(* IEC 61131-3 sources: llm-plc-st-eval/data/processed_definitivo/gpt-4o-2024-08-06/A4/few_shot, 3 files *)

(* ---- ejec_1.st ---- *)
FUNCTION_BLOCK FB_Rampa
VAR_INPUT
    SPvel : REAL; (* Consigna de velocidad *)
    paroRapido : BOOL; (* Activar paro rápido *)
    ciclo : TIME; (* Período de ejecución del bloque *)
END_VAR
VAR_OUTPUT
    CVvel : REAL; (* Velocidad de consigna con rampa *)
END_VAR
VAR
    incremento : REAL; (* Incremento calculado por ciclo *)
    tiempoSegundos : REAL; (* Tiempo de ciclo en segundos *)
END_VAR

(* Convertir el tiempo de ciclo a segundos *)
tiempoSegundos := REAL_TO_REAL(TIME_TO_REAL(ciclo)) / 1000.0;

IF paroRapido THEN
    (* Paro rápido: disminuir CVvel hacia 0.0 con pendiente de 40.0 puntos porcentuales por segundo *)
    incremento := -40.0 * tiempoSegundos;
    CVvel := CVvel + incremento;
    IF CVvel < 0.0 THEN
        CVvel := 0.0;
    END_IF
ELSE
    (* Ajuste normal de CVvel hacia SPvel *)
    IF SPvel > CVvel THEN
        (* Aumentar CVvel hacia SPvel con pendiente de 10.0 puntos porcentuales por segundo *)
        incremento := 10.0 * tiempoSegundos;
        CVvel := CVvel + incremento;
        IF CVvel > SPvel THEN
            CVvel := SPvel;
        END_IF
    ELSIF SPvel < CVvel THEN
        (* Disminuir CVvel hacia SPvel con pendiente de 20.0 puntos porcentuales por segundo *)
        incremento := -20.0 * tiempoSegundos;
        CVvel := CVvel + incremento;
        IF CVvel < SPvel THEN
            CVvel := SPvel;
        END_IF
    END_IF
END_IF
END_FUNCTION_BLOCK

(* ---- ejec_2.st ---- *)
FUNCTION_BLOCK FB_Rampa
VAR_INPUT
    SPvel : REAL; (* Consigna de velocidad *)
    paroRapido : BOOL; (* Señal de paro rápido *)
    ciclo : TIME; (* Período de ejecución del bloque *)
END_VAR
VAR_OUTPUT
    CVvel : REAL; (* Velocidad de consigna con rampa *)
END_VAR
VAR
    incremento : REAL; (* Incremento de velocidad por ciclo *)
    tiempoSegundos : REAL; (* Duración del ciclo en segundos *)
END_VAR

(* Convertir el tiempo de ciclo a segundos *)
tiempoSegundos := REAL_TO_REAL(TIME_TO_REAL(ciclo)) / 1000.0;

IF paroRapido THEN
    (* Paro rápido: disminuir CVvel a 0.0 con pendiente de 40.0 %/s *)
    incremento := -40.0 * tiempoSegundos;
    CVvel := CVvel + incremento;
    IF CVvel < 0.0 THEN
        CVvel := 0.0;
    END_IF
ELSE
    (* Rampa normal: ajustar CVvel hacia SPvel *)
    IF SPvel > CVvel THEN
        (* Incremento al subir con pendiente de 10.0 %/s *)
        incremento := 10.0 * tiempoSegundos;
        CVvel := CVvel + incremento;
        IF CVvel > SPvel THEN
            CVvel := SPvel;
        END_IF
    ELSIF SPvel < CVvel THEN
        (* Decremento al bajar con pendiente de 20.0 %/s *)
        incremento := -20.0 * tiempoSegundos;
        CVvel := CVvel + incremento;
        IF CVvel < SPvel THEN
            CVvel := SPvel;
        END_IF
    END_IF
END_IF
END_FUNCTION_BLOCK

(* ---- ejec_3.st ---- *)
FUNCTION_BLOCK FB_Rampa
VAR_INPUT
    SPvel : REAL; (* Consigna de velocidad *)
    paroRapido : BOOL; (* Señal de paro rápido *)
    ciclo : TIME; (* Período de ejecución del bloque *)
END_VAR
VAR_OUTPUT
    CVvel : REAL; (* Velocidad de consigna con rampa *)
END_VAR
VAR
    deltaTiempo : REAL; (* Tiempo de ciclo en segundos *)
    incremento : REAL; (* Incremento de velocidad por ciclo *)
END_VAR

(* Convertir el tiempo de ciclo a segundos *)
deltaTiempo := REAL_TO_REAL(TIME_TO_REAL(ciclo)) / 1000.0;

IF paroRapido THEN
    (* Paro rápido: descender a 0.0 con pendiente de 40.0 %/s *)
    incremento := -40.0 * deltaTiempo;
    CVvel := CVvel + incremento;
    IF CVvel < 0.0 THEN
        CVvel := 0.0;
    END_IF
ELSE
    (* Ajuste normal de velocidad con rampa *)
    IF SPvel > CVvel THEN
        (* Incremento al subir: máximo 10.0 %/s *)
        incremento := 10.0 * deltaTiempo;
        CVvel := CVvel + incremento;
        IF CVvel > SPvel THEN
            CVvel := SPvel;
        END_IF
    ELSIF SPvel < CVvel THEN
        (* Decremento al bajar: máximo 20.0 %/s *)
        incremento := -20.0 * deltaTiempo;
        CVvel := CVvel + incremento;
        IF CVvel < SPvel THEN
            CVvel := SPvel;
        END_IF
    END_IF
END_IF
END_FUNCTION_BLOCK
